Staubli VAL3: main.pgx

program main()
begin
  close(tCurrentTool)
  pPointRs.config.shoulder = lefty
  pPointRs2.config.shoulder = lefty
  mCurrentSpeed.tvel = 100.00
  mCurrentSpeed.blend = joint
  mCurrentSpeed.reach = 0.010
  mCurrentSpeed.leave = 0.010
  // Program SetProg start
  // Program generated by RoboDK v6.0.7 for Staubli TP80 on XX/XX/XXXX 18:00:00
  // Using nominal kinematics.
  call MoveJoint(10.00000,-20.00000,50.00000,30.00000)
  // Linear movement using joint targets is not supported. Change the target type to cartesian or use a joint movement.
  // Circular movement using joint targets is not supported. Change the target type to cartesian or use a joint movement.
  call MoveJoint(30.00000,25.00000,80.00000,-45.00000)
  delay(0.250)
  call MoveJoint(30.00000,-20.00000,40.00000,60.00000)

  waitEndMove()
  // Program SetProg end

end
